(* IEC 61131-3 sources: 2026_Projet_YGO_ExcavatriceDragage/CODE/J_SUPERVISION/_TYPES/3_CYCLE_ET_MODES, 19 files *)

(* ---- E_CycleDepthStopMode.st ---- *)
(* Mode d'arret de la recherche fond AX7. *)
TYPE E_CycleDepthStopMode :
(
    KOBOLD_ONLY       := 0, // Comportement historique : fond valide par DI Kobold
    SETPOINT_ONLY     := 1, // Arret sur consigne de profondeur valide
    KOBOLD_OR_SETPOINT:= 2  // Premier evenement valide des deux
);
END_TYPE

(* ---- E_CycleSampleCountResetMode.st ---- *)
(* Mode de remise a zero AUTOMATIQUE du compteur JOURNALIER de prelevements.
   Reglage IHM persistant : le comportement se choisit par parametrage, sans modifier le code.
   ⚠️ Le compteur TOTALISATEUR (_CycleSampleCountTotal) n'est JAMAIS concerne par ce
   reglage : aucun mode ne l'ecrit, aucun chemin de RAZ n'existe pour lui.
   🔒 Repli sur valeur non reconnue (memoire persistante restauree hors plage, saisie IHM
   invalide) : aucun des deux modes n'est alors reconnu, donc AUCUNE RAZ automatique ->
   comportement NEVER, le plus conservateur. Le compteur journalier ne peut pas etre efface
   par accident. *)
TYPE E_CycleSampleCountResetMode :
(
    NEVER              := 0, // Defaut : RAZ manuelle IHM uniquement (comportement historique, aucun changement)
    ON_FIRST_START     := 1, // RAZ au premier demarrage de cycle apres mise sous tension de l'automate
    ON_SAFETY_REARM    := 2  // RAZ au rearmement de la chaine AU (contacteur puissance reengage)
);
END_TYPE

(* ---- E_ProgramSequence.st ---- *)
(* =======================================================================
   🔄 E_ProgramSequence — Énumération des séquences de programme automatiques
   ───────────────────────────────────────────────────────────────
   🎯 Rôle : Identifie la séquence active arbitree dans PRG_03
   📄 Référentiel : DOC/WFLOW/CONTRACTS/INTERPRG_CONTRACT_PRG03_MODES_CYCLE_v1.0.md
   ======================================================================= *)
TYPE E_ProgramSequence :
(
    NONE        := 0, // Aucune séquence active
    MAIN_CYCLE  := 1, // Cycle semi-automatique principal (FB_Cycle)
    DIVE_SEARCH := 2, // Recherche de fond Kobold (réservé future migration)
    EXTRACTION  := 3  // Séquence d'extraction (réservé future migration)
);
END_TYPE

(* ---- ST_ChainCycleSemiAuto.st ---- *)
(* =======================================================================
   🔄 ST_ChainCycleSemiAuto — Diagnostic chronologique Séquenceur Semi-Auto
   ───────────────────────────────────────────────────────────────
   🎯 Rôle : Vue dépannage / Watch CODESYS pour le cycle semi-automatique
   📄 Doc métier : DOC/AF/AF_Partie-14_Fonction_Troubleshooting/FB_TroubleshootingView_v1.2.md
   🔒 Sécurité : 100% lecture seule / diagnostic d'observation
   ======================================================================= *)

TYPE ST_ChainCycleSemiAuto :
STRUCT
    // 🚦 1. Conditions d'engagement et autorisations
    Idx101_ModeSemiAutoActive        : BOOL; // 1 = Mode arbitré SEMI_AUTO actif | 0 = Autre mode
    Idx102_PowerAndSafetyOk          : BOOL; // 1 = Chaîne de sécurité OK (PowerContactorEngaged)
    Idx103_HeartbeatIhmOk            : BOOL; // 1 = Liaison IHM<->PLC valide
    Idx104_DeadmanArmed              : BOOL; // 1 = Bouton homme-mort armé (fenêtre 3s active)
    Idx105_MancheDeflechi            : BOOL; // 1 = Permis mouvement armé (manche hors zone neutre)
    Idx106_HomedM1M2                 : BOOL; // 1 = Codeurs treuils M1 et M2 référencés
    Idx107_StartCycleRequest         : BOOL; // 1 = Demande Start reçue (IHM)
    Idx108_AbortCycleRequest         : BOOL; // 1 = Demande Abort reçue (IHM)

    // 🔄 2. État du Séquenceur
    Idx201_Ready                     : BOOL; // 1 = Séquenceur prêt à démarrer
    Idx202_Busy                      : BOOL; // 1 = Cycle en cours d'exécution
    Idx203_Done                      : BOOL; // 1 = Cycle terminé avec succès
    Idx204_Error                     : BOOL; // 1 = Défaut vue LIVE (retombe seul avec la cause)
    Idx205_ErrorId                   : WORD; // Code d'erreur interne FB_Cycle
    Idx217_FaultLatched              : BOOL; // 1 = Défaut vue LATCHÉE (bloque AX0->AX1 même si Idx204=0, exige Reset conscient)
    Idx218_FaultLatchedId            : WORD; // Bitfield fige a l'apparition du defaut latche
    Idx219_CycleChecksInhibited       : BOOL; // 1 = controles procede inhibes, protections actives
    Idx220_IgnoredCycleCheckId        : WORD; // Causes procede actives mais ignorees
    // ⚠️ Idx221 (ForceStepPrepared) SUPPRIME par T358 : le mecanisme a deux temps du
    //    forcage de step n'existe plus (saut immediat sans preparation). L'index reste
    //    VACANT pour ne renumeroter aucun tag IHM de la chaine de depannage.
    Idx222_ForceStepResult            : STRING(120); // Motif de rejet de la derniere consigne de forcage (T358)
    Idx206_Step                      : E_AutoCycleStep; // Étape courante (X0 à X13 + AX_STAB)
    Idx207_StepStr                   : STRING(80);  // Libellé explicite de l'étape
    Idx208_StepAtError               : E_AutoCycleStep; // Étape mémorisée lors du dernier défaut
    Idx209_WaitingForOperator        : BOOL;        // 1 = En attente d'une action humaine
    Idx210_WaitingForProcess         : BOOL;        // 1 = En attente d'une condition physique/procédé
    Idx211_OperatorActionId          : WORD;        // Identifiant numérique de l'action attendue
    Idx212_OperatorAction            : STRING(120); // Description explicite de l'action/attente
    Idx213_ExpectedAxis              : E_OperatorAxis; // Organe attendu (NONE, JOYSTICK_X, JOYSTICK_Y, BUTTON)
    Idx214_ExpectedDirection         : INT;         // Sens attendu (-1, 0, +1)
    Idx215_WaitingResume             : BOOL;        // 1 = En pause suite à bascule de mode (attente StartCycle)
    Idx216_PausedState               : E_AutoCycleStep; // Étape mémorisée prête pour reprise

    // 🎯 3. Consignes & Feedbacks Opérationnels
    Idx301_TargetPosition            : INT;  // Cible translation sélectionnée (1=Trémie, 3=P1)
    Idx302_TargetDepth_M             : REAL; // Profondeur de consigne (m)
    Idx303_KoboldBottomTouch         : BOOL; // 1 = Détection contact fond Kobold
    Idx304_SpeedMismatchActive       : BOOL; // 1 = Alerte écart de vitesse M1/M2 active
    Idx305_LimitLegalReached         : BOOL; // 1 = Limite légale atteinte (descente bloquée)
    Idx306_WinchSyncError            : BOOL; // 1 = Erreur de synchronisme M1/M2
    Idx307_M1SpeedStepApplied        : INT;  // Palier vitesse applique M1 (0..5, causes 8/9)
    Idx308_M2SpeedStepApplied        : INT;  // Palier vitesse applique M2 (0..5, causes 8/9)
    Idx309_AutoDiveM2Step5Active     : BOOL; // 1 = Essai T291-A actif (M2 cible palier 5 en plongee)
    Idx310_M1SpeedStepAtFault        : INT;  // Palier M1 applique, fige au moment du defaut (0..5)
    Idx311_M2SpeedStepAtFault        : INT;  // Palier M2 applique, fige au moment du defaut (0..5)
END_STRUCT
END_TYPE

(* ---- ST_CycleCmd.st ---- *)
(* ═══════════════════════════════════════════════════════════════
   🎮 ST_CycleCmd — Commandes IHM pour le cycle semi-automatique
   ═══════════════════════════════════════════════════════════════ *)
TYPE ST_CycleCmd :
STRUCT
    BtnStart          : BOOL; (* ▶️ Lancement cycle automatique *)
    BtnPause          : BOOL; (* ⏸️ Pause cycle automatique *)
    BtnAbort          : BOOL; (* ⏹️ Abandon / arrêt cycle automatique *)
    BtnResumeAfterFault : BOOL; (* Reprise consciente depuis AX_STAB vers l'etape d'origine *)
    BtnReset          : BOOL; (* 🔁 Reset dédié FB_Cycle, jamais mélangé au reset défauts général () *)
    BtnSkipDrain      : BOOL; (* ⏭️ Passer l'étape d'égouttage X9 (front) *)
    BtnReposition     : BOOL; (* ⬇️ Option maintenue : repositionnement couplé M1+M2 pendant le vidage trémie (X11b <-> X11c) *)
    TglCommissioning  : BOOL := FALSE; (* 🔧 Case mise en service : déverrouille le forçage de step (front/impulsion). NON persisté. *)
    TglCycleChecksInhibit : BOOL := FALSE; (* 🧪 Mode essai : inhibe uniquement les controles procede autorises. NON persiste. *)
    TglAutoDiveM2Step5Trial : BOOL := TRUE; (* Profil nominal : en SEMI_AUTO AX4..AX7, M1 reste palier 4 et M2 peut monter au palier 5. Debrayable IHM, non persiste. *)
    BtnResetSampleCount : BOOL; (* 🔢 RAZ consciente du compteur JOURNALIER de prélèvements (front) — n'agit JAMAIS sur le totalisateur, qui n'a aucune commande *)
    // ⚠️ AJOUT EN FIN DE STRUCT (mapping positionnel : jamais d'insertion au milieu).
    // 🔧 T358 : consigne de forcage de step — VALEUR écrite par l'opérateur, lue ET
    //    acquittee par FB_CycleSemiAuto (retour à la sentinelle -1). Remplace le couple
    //    BtnForceStepApply + ST_CycleCfg.ForceStepTarget : plus de bouton, plus de
    //    confirmation, plus de cible persistée (donc aucun saut d'étape au démarrage).
    //    Zone Cmd = NON persistée : la consigne ne survit jamais à une coupure.
    //    -1 = aucune demande ; 0..22 = étape cible (plage E_AutoCycleStep).
    SetForceStepTgt : INT := -1; (* 🔧 Étape cible du forçage immédiat du cycle ; -1 = aucune demande *)
    // Options souplesse cycle vidage tremie & conditions initiales (non persistees, zero decalage GVL_PERSISTENT)
    TglAllowDumpInPV      : BOOL := FALSE; (* 🪣 Autorise l'ouverture benne dès la zone PV + retour P1 dès benne ouverte sans exiger capteur Trémie *)
    TglRelaxSemiAutoStart : BOOL := FALSE; (* 🟢 Assouplit les conditions initiales en AX1_INIT (fenêtre haute élargie + dispense qualification benne si treuils hauts) *)
    SetPauseBeforeDump_S  : REAL := 0.0;   (* ⏱️ Pause réglable (s) entre l'arrêt translation AX14 et l'ouverture benne AX15B (0.0 = transparent) *)
END_STRUCT
END_TYPE

(* ---- ST_CycleHMI.st ---- *)
(* ═══════════════════════════════════════════════════════════════
   🔄 ST_CycleHMI — Données d'échange IHM du cycle semi-automatique
   ───────────────────────────────────────────────────────────────
   📄 Structuration en Cmd / State / Cfg / Test , homogène avec ST_WinchHMI.
   Cfg protégé par persistance GVL_PERSISTENT
   ═══════════════════════════════════════════════════════════════ *)
TYPE ST_CycleHMI :
STRUCT
    Cmd   : ST_CycleCmd;
    State : ST_CycleState;
    Cfg   : ST_CycleCfg;
END_STRUCT
END_TYPE

(* ---- ST_CycleMachineHomingCfg.st ---- *)
(* ═══════════════════════════════════════════════════════════════
   ⚙️ ST_CycleMachineHomingCfg — Réglages IHM du cycle de référencement machine
   ───────────────────────────────────────────────────────────────
   🎯 Mise en service. Les réglages géométriques (positions capteur, offsets benne)
      restent portés par GVL_PERSISTENT (_WinchM1CfgPersist / _BucketCfgPersist).
   💾 Ponté vers persist (_CycleMachineHomingCfgPersist) via FB_CfgPersistBridge_CycleMachineHomingCfg.
   ═══════════════════════════════════════════════════════════════ *)
TYPE ST_CycleMachineHomingCfg :
STRUCT
    ForceStepTarget : INT  := 0;     (* 🔧 Step GRAFCET cible du forçage (0=HX0 .. 9=HXF), borné côté FB *)
    Initialized     : BOOL := FALSE; (* 🚦 flag restauration boot *)
END_STRUCT
END_TYPE

(* ---- ST_CycleMachineHomingCmd.st ---- *)
(* ═══════════════════════════════════════════════════════════════
   🎮 ST_CycleMachineHomingCmd — Commandes IHM du cycle de référencement machine
   ───────────────────────────────────────────────────────────────
   🎯 Cycle homing machine (FB_CycleMachineHoming) — orchestré en MAINT_N2.
      Séparé de ST_CycleCmd (cycle SEMI_AUTO) et de ST_ModesCmd (modes de marche).
      Boutons momentanés uniquement ; réglages -> ST_CycleMachineHomingCfg.
   ═══════════════════════════════════════════════════════════════ *)
TYPE ST_CycleMachineHomingCmd :
STRUCT
    BtnStart          : BOOL; (* ▶️ Lancer le cycle de homing machine (MAINT_N2, front) — alternative au motif 3 appuis joystick *)
    BtnValidate       : BOOL; (* ✅ Validation depuis IHM (front) — équivaut à 1 appui du motif 3 appuis joystick *)
    BtnAbort          : BOOL; (* ⏹️ Quitter / abandonner le cycle homing (front) — retour HX0 sans mouvement *)
    TglCommissioning  : BOOL := FALSE; (* 🔧 Case mise en service : déverrouille le forçage de step (MAINT_N2). NON persisté (reset au reboot = sûr). *)
    BtnForceStepApply : BOOL; (* 🔧 Applique le forçage de step (front) — impulsion ; cible = ST_CycleMachineHomingCfg.ForceStepTarget *)
END_STRUCT
END_TYPE

(* ---- ST_CycleMachineHomingHMI.st ---- *)
(* ═══════════════════════════════════════════════════════════════
   🎯 ST_CycleMachineHomingHMI — Données d'échange IHM du cycle de référencement machine
   ───────────────────────────────────────────────────────────────
   📄 Structuration Cmd / State / Cfg , homogène avec ST_CycleHMI /
      ST_CycleDiveSearchHMI / ST_CycleExtractionHMI.
   ═══════════════════════════════════════════════════════════════ *)
TYPE ST_CycleMachineHomingHMI :
STRUCT
    Cmd   : ST_CycleMachineHomingCmd;
    State : ST_MachineHoming;      (* Image publiée du FB_CycleMachineHoming (SeqStep, Step, Instruction, Failed, ordres, …) *)
    Cfg   : ST_CycleMachineHomingCfg;
END_STRUCT
END_TYPE

(* ---- ST_MaintenanceN2HMI.st ---- *)
(* ═══════════════════════════════════════════════════════════════
   🛠️ ST_MaintenanceN2HMI — Données d'échange IHM pour la maintenance N2
   ───────────────────────────────────────────────────────────────
   📄 Structuration canonique Cmd / State pour la maintenance experte N2.
   ═══════════════════════════════════════════════════════════════ *)
TYPE ST_MaintenanceN2HMI :
STRUCT
    Cmd   : ST_MaintenanceN2Cmd;
    State : ST_MaintenanceN2State;
END_STRUCT
END_TYPE

(* ---- ST_Modes_Autorisations.st ---- *)
(* =======================================================================
   ST_Modes_Autorisations - Bus public d'autorisations du mode machine
   -----------------------------------------------------------------------
   Doc metier : DOC/AF/AF_Partie-05_Modes_Maintenance_v2.1.md
                DOC/AF/AF_Partie-02_Architecture_Programme_v3.2.md #2
   NC-110 : le prefixe ST_fb* est reserve aux DUT propriete d'un seul FB.
      Ce DUT est un BUS multi-consommateurs (>=6 domaines : Cycle, Safety,
      Treuils, Translation, Supervision, Acquisition) -> renomme
      ST_Modes_Autorisations (bus de domaine public, sans le prefixe FB).
   Produit par FB_Modes (via PRG_03_Modes_Cycle)
      Consomme par : Cycle, Safety, Treuils, Translation, Supervision, Acquisition
   Producteur unique : FB_Modes (via PRG_03_Modes_Cycle)
   ======================================================================= *)

TYPE ST_Modes_Autorisations :
STRUCT
    Mode                        : E_Mode;     // Mode arbitre (DISABLE/N1/N2/SEMI_AUTO)
    SyncEnable                  : BOOL;       // Synchro M1/M2 (logique positive)
    InhibitM1                   : BOOL;       // Inhibition M1 (MAINT_N2 only)
    InhibitM2                   : BOOL;       // Inhibition M2 (MAINT_N2 only)
    JoystickWinchSelectArbitrated : INT;      // 0=M1+M2 couples nominal, 1=M1, 2=M2 (unitaires MAINT_N2)
    CoupledBucketPhaseLocked    : BOOL;       // T248 : phase mouvement couple VERROUILLEE pour ce maintien joystick -> la perte de l'etat ouvert/ferme en mouvement ne relance PAS de correction benne, ni de blocage "descente/montee interdite". Efface au relachement joystick confirme.
    WinchSelTransitionHold      : BOOL;       // T248 : changement de selecteur en cours -> requetes mouvement M1/M2 forcees a 0 jusqu'a l'arret confirme (pas de hand-off en mouvement)
    HomingApproachEnable        : BOOL;       // Depassement butee haut (N2)
    MaintenanceM3TargetEnable   : BOOL;       // Cible Translation Maintenance (N2 only)

    // AF-05 #4bis - matrice de maintenance
    // Ces trois champs sont des FAITS/DIAGS publies, pas des autorisations : ils
    // restent vrais meme quand le FB est neutralise par Enable=FALSE (etat persistant).
    ModeChangePendingBlocked    : BOOL;       // Demande de changement de mode REFUSEE : les treuils
                                              //   ne sont pas a l'arret mecanique confirme (contacteurs
                                              //   retombes ET frein serre ET |v| < seuil). Mode courant maintenu.
    ModeChangeBlockReason       : STRING(40); // Motif du blocage de bascule (texte IHM court, ex. "Chgt mode refuse : contacteur M1")
    // Détail des 6 sous-conditions de ModeChangeAllowed (diagnostic IHM) — TRUE = condition satisfaite.
    M1ContactorsReleased        : BOOL;       // M1 : contacteurs retombés
    M1BrakeApplied              : BOOL;       // M1 : frein serré (NOT M1BrakeIsOpen)
    M1SpeedLow                  : BOOL;       // M1 : vitesse sous seuil
    M2ContactorsReleased        : BOOL;       // M2 : contacteurs retombés
    M2BrakeApplied              : BOOL;       // M2 : frein serré (NOT M2BrakeIsOpen)
    M2SpeedLow                  : BOOL;       // M2 : vitesse sous seuil
    HomingRequiredM1            : BOOL;       // M1 : re-homing obligatoire avant tout retour SEMI_AUTO
    HomingRequiredM2            : BOOL;       // M2 : idem
END_STRUCT
END_TYPE

(* ---- ST_ModesCycleInterPrg.st ---- *)
(* =======================================================================
   📦 ST_ModesCycleInterPrg — Bus public d'autorisations et demandes de cycle
   ───────────────────────────────────────────────────────────────
   🎯 Rôle : Structure de données globale publiée par PRG_03_Modes_Cycle
   📄 Référentiel : DOC/WFLOW/CONTRACTS/INTERPRG_CONTRACT_PRG03_MODES_CYCLE_v1.0.md
   ======================================================================= *)
TYPE ST_ModesCycleInterPrg :
STRUCT
    Auth          : ST_Modes_Autorisations; // Bus public d'autorisations machine (NC-110)
    WinchBothIntent : ST_WinchBothIntent;     // 🎮 Intention both continue opérateur (source unique PRG_03, TOUS modes)
    AutoDiveM1Step4M2Step5Active : BOOL;      // Essai T291-A actif : SEMI_AUTO AX4..AX7, descente M1 palier 4 / M2 palier 5
    ReqProgram    : ST_ProgramRequest;        // Demandes programme vers PRG_04 / PRG_05
    SequenceState : ST_SequencePublicState;   // État public de la séquence
    // 🧩 Défaut de l'arbitre de mode (FB_Modes), forme cible ST_Fault (AF03 §3).
    // Producteur unique : FB_Modes (instancié par PRG_03_Modes_Cycle).
    // Causes : [0] refus Semi-Auto pour défaut codeur (latchée) ;
    //          [1] changement de mode refusé, treuils non à l'arrêt confirmé (live) ;
    //          [2] refus Semi-Auto pour re-homing obligatoire (latchée).
    // ⚠️ Sans cette publication, les refus de mode restaient invisibles de l'IHM :
    //    un interlock qu'on ne voit pas est un interlock qu'on contourne.
    ModesFault    : ST_Fault;                 // 🚨 Défauts d'arbitrage de mode (consommé PRG_07 → IHM)
END_STRUCT
END_TYPE

(* ---- ST_ModesHMI.st ---- *)
(* ═══════════════════════════════════════════════════════════════
   🎚️ ST_ModesHMI — Données d'échange IHM pour les modes de marche
   ───────────────────────────────────────────────────────────────
   📄 Structuration en Cmd / State , homogène avec ST_WinchHMI/ST_SyncHMI/ST_BucketHMI.
   Pas de Cfg (aucun réglage numérique dans ce domaine) ni de Bypass (concept absent de Modes).
   ═══════════════════════════════════════════════════════════════ *)
TYPE ST_ModesHMI :
STRUCT
    Cmd   : ST_ModesCmd;
    State : ST_ModesState;
END_STRUCT
END_TYPE

(* ---- ST_ModesState.st ---- *)
(* ═══════════════════════════════════════════════════════════════
   🚦 ST_ModesState — États et diagnostics IHM des modes de marche
   ═══════════════════════════════════════════════════════════════ *)
TYPE ST_ModesState :
STRUCT
    CurrentMode           : E_Mode; (* 🎚️ Mode de marche actuellement actif *)
    AnyFaultActive        : BOOL;   (* : au moins un défaut/alarme actif dans le domaine
                                        sécurité/métier — s'éteint seul quand la cause disparaît ET que
                                        BtnFaultReset a été pressé (OR de tous les .Error du domaine,
                                        même périmètre que BtnFaultReset) *)

    (* Miroir IHM des états de maintenance (AF-05 §4bis) *)
    ModeChangePendingBlocked : BOOL;   (* 🚦 Changement de mode refusé : treuils non à l'arrêt confirmé (contacteurs retombés + frein serré + |v| < seuil) *)
    ModeChangeBlockReason    : STRING(40); (* 🚦 Motif du blocage de bascule (texte court, ex. "Chgt mode refuse : contacteur M1") *)
    (* Détail des 6 sous-conditions de ModeChangeAllowed (diagnostic IHM) — TRUE = condition satisfaite *)
    M1ContactorsReleased : BOOL; (* M1 : contacteurs retombés *)
    M1BrakeApplied       : BOOL; (* M1 : frein serré *)
    M1SpeedLow           : BOOL; (* M1 : vitesse sous seuil *)
    M2ContactorsReleased : BOOL; (* M2 : contacteurs retombés *)
    M2BrakeApplied       : BOOL; (* M2 : frein serré *)
    M2SpeedLow           : BOOL; (* M2 : vitesse sous seuil *)
    HomingRequiredM1         : BOOL;   (* 🧭 M1 : re-homing obligatoire avant retour SEMI_AUTO *)
    HomingRequiredM2         : BOOL;   (* 🧭 M2 : re-homing obligatoire avant retour SEMI_AUTO *)
END_STRUCT
END_TYPE

(* ---- ST_OperatorCoupledIntent.st ---- *)
(* =======================================================================
   🎮 ST_WinchBothIntent — Intention both continue de l'opérateur
   ───────────────────────────────────────────────────────────────
   🎯 Rôle : Transmet l'intention de mouvement both (2 treuils ensemble,
      homme-mort / boutons) produite inconditionnellement par PRG_03 vers
      PRG_04 et l'arbitrage (tous modes). Source UNIQUE de la décision both.
   📄 Référentiel : DOC/WFLOW/CONTRACTS/INTERPRG_CONTRACT_PRG03_MODES_CYCLE_v1.0.md
   ======================================================================= *)
TYPE ST_WinchBothIntent :
STRUCT
    Active      : BOOL; // Intention both active (homme-mort qualifié + Select=0 OU boutons BothUp/BothDown)
    ReqAscent   : BOOL; // Intention both montée
    ReqDescend  : BOOL; // Intention both descente
END_STRUCT
END_TYPE

(* ---- ST_ProgramBucketRequest.st ---- *)
(* =======================================================================
   🪣 ST_ProgramBucketRequest — Demande de mouvement benne par le programme
   ───────────────────────────────────────────────────────────────
   🎯 Rôle : Regroupe les demandes logiques de manœuvre benne et mesure Kobold
   📄 Référentiel : DOC/WFLOW/CONTRACTS/INTERPRG_CONTRACT_PRG03_MODES_CYCLE_v1.0.md
   ======================================================================= *)
TYPE ST_ProgramBucketRequest :
STRUCT
    ReqOpen                     : BOOL; // Demande ouverture benne
    ReqClose                    : BOOL; // Demande fermeture benne
    ReqHoldAscentP1AfterClose   : BOOL; // Maintien M2 en montee P1 apres fermeture, pour raccordement AX10B sans coupure
    ReqKoboldMeasureEnable      : BOOL; // Demande activation mesure/contacteur Kobold
    DescendPermitDiveBucketOpen : BOOL; // Autorisation de descente conditionnée benne ouverte (DiveSearch)
    ExtractionControlActive     : BOOL; // Plafond palier 1 pendant la montée contrôlée
    AscentPermit                : BOOL; // Autorisation de remontée assistée (ExtractionAssist)
    MinStepDown                 : INT;  // Palier plancher de descente imposé pendant la plongée (FB_DiveSearch, 0 = aucun)
END_STRUCT
END_TYPE

(* ---- ST_ProgramRequest.st ---- *)
(* =======================================================================
   📋 ST_ProgramRequest — Ensemble des demandes de mouvements du programme
   ───────────────────────────────────────────────────────────────
   🎯 Rôle : Regroupe les demandes formulées vers PRG_04 (Treuils/Benne) et PRG_05 (Translation)
   📄 Référentiel : DOC/WFLOW/CONTRACTS/INTERPRG_CONTRACT_PRG03_MODES_CYCLE_v1.0.md
   ======================================================================= *)
TYPE ST_ProgramRequest :
STRUCT
    ReqWinchM1            : ST_ProgramWinchRequest;       // Demande programme treuil M1
    ReqWinchM2            : ST_ProgramWinchRequest;       // Demande programme treuil M2
    ReqTranslation        : ST_ProgramTranslationRequest; // Demande programme translation M3
    ReqBucket             : ST_ProgramBucketRequest;      // Demande programme benne
END_STRUCT
END_TYPE

(* ---- ST_ProgramTranslationRequest.st ---- *)
(* =======================================================================
   🎯 ST_ProgramTranslationRequest — Demande de mouvement translation par le programme
   ───────────────────────────────────────────────────────────────
   🎯 Rôle : Regroupe les demandes logiques de translation M3 formulées par le séquenceur
   📄 Référentiel : DOC/WFLOW/CONTRACTS/INTERPRG_CONTRACT_PRG03_MODES_CYCLE_v1.0.md
   ======================================================================= *)
TYPE ST_ProgramTranslationRequest :
STRUCT
    ReqStart    : BOOL; // Demande de démarrage mouvement translation
    PositionTgt : INT;  // Cible de position demandée (1=Trémie, 2=P2, 3=P1, 4=Maintenance)
END_STRUCT
END_TYPE

(* ---- ST_ProgramWinchRequest.st ---- *)
(* =======================================================================
   🔌 ST_ProgramWinchRequest — Demande de mouvement treuil par le programme
   ───────────────────────────────────────────────────────────────
   🎯 Rôle : Regroupe les demandes logiques de treuil formulées par le séquenceur
   📄 Référentiel : DOC/WFLOW/CONTRACTS/INTERPRG_CONTRACT_PRG03_MODES_CYCLE_v1.0.md
   ======================================================================= *)
TYPE ST_ProgramWinchRequest :
STRUCT
    RunRequest   : BOOL; // Ordre marche demandé par le programme
    ReqAscent    : BOOL; // Demande montée
    ReqDescend   : BOOL; // Demande descente
    StepTgt      : INT;  // Palier de vitesse cible demandé (1 à 5, 0 = arrêt)
END_STRUCT
END_TYPE
